(* IEC 61131-3 sources: plc-iiot-stack/tests/POUs/FB_MqttClientFake, 22 files *)

(* ---- FB_MqttClientFake.decl.st ---- *)
// Назначение: подменный клиент MQTT для тестов (I_MqttClient): связь, отказы подключения, подписки и
//             публикации задаются входами; опубликованные сообщения сохраняются (aPub; фильтр aCapture —
//             только нужные топики), входящие ставятся в очередь методом Inject. Методы поиска по топику
//             безопасны для пустого журнала.
// Автор:      kr0nsch
// Версия:     0.1.0
// Документ:   docs/TEST_REPORT.md
FUNCTION_BLOCK FB_MqttClientFake IMPLEMENTS I_MqttClient
VAR_INPUT
    xLinkUp : BOOL := TRUE;            // брокер доступен: после Connect связь есть сразу
    xConnectAccepts : BOOL := TRUE;    // Connect() возвращает TRUE
    xSubscribeAccepts : BOOL := TRUE;
    xPublishAccepts : BOOL := TRUE;    // FALSE — «очередь полна»
    diError : DINT;                    // значение LastError()
    aCapture : ARRAY[1..CAPTURE_MAX] OF STRING(GVL_Const.MQTT_TOPIC_LEN);   // не пусто — сохранять только эти
END_VAR
VAR_OUTPUT
    xConnectRequested : BOOL;
    uiConnectCalls : UINT;
    uiDisconnectCalls : UINT;
    uiServiceCalls : UINT;
    uiSubscribeCalls : UINT;
    stLastCfg : ST_MqttBrokerCfg;
    sLastFilter : STRING(GVL_Const.MQTT_TOPIC_LEN);
    eLastFilterQos : E_MqttQos;
    uiPubCount : UINT;                 // сообщений в aPub
    uiPubTotal : UINT;                 // принятых публикаций всего (сохранённых и нет)
    uiPubRejected : UINT;              // Publish вернул FALSE
    aPub : ARRAY[1..PUB_MAX] OF ST_FakeMqttMsg;
    uiInCount : UINT;                  // входящих в очереди
END_VAR
VAR
    aIn : ARRAY[1..IN_MAX] OF ST_FakeMqttIn;
END_VAR
VAR CONSTANT
    PUB_MAX : UINT := 48;
    IN_MAX : UINT := 16;
    CAPTURE_MAX : UINT := 8;
END_VAR

(* ---- Captured.method.decl.st ---- *)
// Сохранять ли сообщение: фильтр aCapture пуст или топик в нём.
METHOD PRIVATE Captured : BOOL
VAR_INPUT
    sTopicIn : STRING(GVL_Const.MQTT_TOPIC_LEN);
END_VAR
VAR
    uiIdx : UINT;
    xAny : BOOL;
END_VAR

(* ---- Captured.method.impl.st ---- *)
FOR uiIdx := 1 TO CAPTURE_MAX DO
    IF LEN(aCapture[uiIdx]) > 0 THEN
        xAny := TRUE;
        IF aCapture[uiIdx] = sTopicIn THEN
            Captured := TRUE;
            RETURN;
        END_IF
    END_IF
END_FOR
Captured := NOT xAny;

(* ---- Connect.method.decl.st ---- *)
// I_MqttClient: запоминает параметры; связь появляется, если xLinkUp.
METHOD Connect : BOOL
VAR_IN_OUT CONSTANT
    // lint:allow STL007 параметр VAR_IN_OUT CONSTANT — ссылка только для чтения, а не константа
    stCfg : ST_MqttBrokerCfg;
END_VAR

(* ---- Connect.method.impl.st ---- *)
uiConnectCalls := uiConnectCalls + 1;
stLastCfg := stCfg;
IF xConnectAccepts THEN
    xConnectRequested := TRUE;
    Connect := TRUE;
END_IF

(* ---- CountTopic.method.decl.st ---- *)
// Для тестов: сколько сообщений с топиком sTopic.
METHOD CountTopic : UINT
VAR_INPUT
    sTopic : STRING(GVL_Const.MQTT_TOPIC_LEN);
END_VAR
VAR
    uiIdx : UINT;
END_VAR

(* ---- CountTopic.method.impl.st ---- *)
FOR uiIdx := 1 TO uiPubCount DO
    IF aPub[uiIdx].sTopic = sTopic THEN
        CountTopic := CountTopic + 1;
    END_IF
END_FOR

(* ---- FindLast.method.decl.st ---- *)
// Для тестов: индекс последнего сообщения с топиком sTopic; нет — 0.
METHOD FindLast : UINT
VAR_INPUT
    sTopic : STRING(GVL_Const.MQTT_TOPIC_LEN);
END_VAR
VAR
    diIdx : DINT;
END_VAR

(* ---- FindLast.method.impl.st ---- *)
FOR diIdx := UINT_TO_DINT(uiPubCount) TO 1 BY -1 DO
    IF aPub[diIdx].sTopic = sTopic THEN
        FindLast := DINT_TO_UINT(diIdx);
        RETURN;
    END_IF
END_FOR

(* ---- Inject.method.decl.st ---- *)
// Для тестов: поставить входящее сообщение в очередь. FALSE — очередь полна.
METHOD Inject : BOOL
VAR_INPUT
    sTopic : STRING(GVL_Const.MQTT_TOPIC_LEN);
    sPayload : STRING(GVL_Const.MQTT_CMD_PAYLOAD_LEN);
    xTruncated : BOOL;
    xRetained : BOOL;
END_VAR

(* ---- Inject.method.impl.st ---- *)
IF uiInCount >= IN_MAX THEN
    RETURN;
END_IF
uiInCount := uiInCount + 1;
aIn[uiInCount].sTopic := sTopic;
aIn[uiInCount].sPayload := sPayload;
aIn[uiInCount].xTruncated := xTruncated;
aIn[uiInCount].xRetained := xRetained;
Inject := TRUE;

(* ---- LastHas.method.decl.st ---- *)
// Для тестов: последнее сообщение с топиком sTopic содержит sPart.
METHOD LastHas : BOOL
VAR_INPUT
    sTopic : STRING(GVL_Const.MQTT_TOPIC_LEN);
    sPart : STRING(255);
END_VAR
VAR
    uiIdx : UINT;
END_VAR

(* ---- LastHas.method.impl.st ---- *)
uiIdx := FindLast(sTopic := sTopic);
IF uiIdx > 0 THEN
    LastHas := F_TestContains(sText := aPub[uiIdx].sPayload, sPart := sPart);
END_IF

(* ---- LastIs.method.decl.st ---- *)
// Для тестов: последнее сообщение с топиком sTopic равно sExpected (до 255 символов).
METHOD LastIs : BOOL
VAR_INPUT
    sTopic : STRING(GVL_Const.MQTT_TOPIC_LEN);
    sExpected : STRING(255);
END_VAR
VAR
    uiIdx : UINT;
END_VAR

(* ---- LastIs.method.impl.st ---- *)
uiIdx := FindLast(sTopic := sTopic);
IF uiIdx > 0 THEN
    LastIs := aPub[uiIdx].sPayload = sExpected;
END_IF

(* ---- LastPayload.method.decl.st ---- *)
// Для тестов: начало (255 символов) последнего сообщения с топиком sTopic — для текста отказа.
METHOD LastPayload : STRING(255)
VAR_INPUT
    sTopic : STRING(GVL_Const.MQTT_TOPIC_LEN);
END_VAR
VAR
    uiIdx : UINT;
END_VAR

(* ---- LastPayload.method.impl.st ---- *)
uiIdx := FindLast(sTopic := sTopic);
IF uiIdx > 0 THEN
    LastPayload := aPub[uiIdx].sPayload;
ELSE
    LastPayload := '<none>';
END_IF

(* ---- Publish.method.decl.st ---- *)
// I_MqttClient: принимает сообщение и сохраняет его в aPub (с учётом фильтра aCapture).
METHOD Publish : BOOL
VAR_INPUT
    sTopic : STRING(GVL_Const.MQTT_TOPIC_LEN);
    eQos : E_MqttQos;
    xRetain : BOOL;
END_VAR
VAR_IN_OUT CONSTANT
    // lint:allow STL007 параметр VAR_IN_OUT CONSTANT — ссылка только для чтения, а не константа
    sPayload : STRING(GVL_Const.MQTT_PAYLOAD_LEN);
END_VAR

(* ---- Publish.method.impl.st ---- *)
IF NOT IsConnected() OR NOT xPublishAccepts THEN
    uiPubRejected := uiPubRejected + 1;
    RETURN;
END_IF
Publish := TRUE;
uiPubTotal := uiPubTotal + 1;
IF NOT Captured(sTopicIn := sTopic) OR uiPubCount >= PUB_MAX THEN
    RETURN;
END_IF
uiPubCount := uiPubCount + 1;
aPub[uiPubCount].sTopic := sTopic;
aPub[uiPubCount].sPayload := sPayload;
aPub[uiPubCount].eQos := eQos;
aPub[uiPubCount].xRetain := xRetain;

(* ---- Receive.method.decl.st ---- *)
// I_MqttClient: первое сообщение очереди входящих.
METHOD Receive : BOOL
VAR_IN_OUT
    sTopic : STRING(GVL_Const.MQTT_TOPIC_LEN);
    sPayload : STRING(GVL_Const.MQTT_CMD_PAYLOAD_LEN);
END_VAR
VAR_OUTPUT
    xTruncated : BOOL;
    xRetained : BOOL;
END_VAR
VAR
    uiIdx : UINT;
END_VAR

(* ---- Receive.method.impl.st ---- *)
IF uiInCount = 0 OR NOT IsConnected() THEN
    RETURN;
END_IF
sTopic := aIn[1].sTopic;
sPayload := aIn[1].sPayload;
xTruncated := aIn[1].xTruncated;
xRetained := aIn[1].xRetained;
FOR uiIdx := 1 TO uiInCount - 1 DO
    aIn[uiIdx] := aIn[uiIdx + 1];
END_FOR
uiInCount := uiInCount - 1;
Receive := TRUE;

(* ---- Subscribe.method.decl.st ---- *)
// I_MqttClient: запоминает фильтр.
METHOD Subscribe : BOOL
VAR_INPUT
    sTopicFilter : STRING(GVL_Const.MQTT_TOPIC_LEN);
    eQos : E_MqttQos;
END_VAR
